Staubli VAL3: _clickIoPage.pgx

public program _clickIoPage()
begin
  sPageUsing="InOut"
  userPage("Disk://source/projectSource/io/interface/InOut")
  delay(1)
end
